(* IEC 61131-3 sources: STruCpp/tests/st-validation/oscat, 20 files *)

(* ---- oscat_bits.st ---- *)
FUNCTION BIT_TOGGLE_B : BYTE
VAR_INPUT
	IN : BYTE;
	POS : INT;
END_VAR
BIT_TOGGLE_B := SHL(BYTE#1, POS) XOR IN;
END_FUNCTION

FUNCTION BYTE_TO_GRAY : BYTE
VAR_INPUT
	IN : BYTE;
END_VAR
BYTE_TO_GRAY := IN XOR SHR(IN,1);
END_FUNCTION

FUNCTION GRAY_TO_BYTE : BYTE
VAR_INPUT
	IN : BYTE;
END_VAR
GRAY_TO_BYTE := SHR(IN,4) XOR IN;
GRAY_TO_BYTE := SHR(GRAY_TO_BYTE,2) XOR GRAY_TO_BYTE;
GRAY_TO_BYTE := SHR(GRAY_TO_BYTE,1) XOR GRAY_TO_BYTE;
END_FUNCTION

(* ---- oscat_convert.st ---- *)
(* OSCAT Conversion Functions — Unit conversions and range mapping *)

FUNCTION KMH_TO_MS : REAL
VAR_INPUT
	KMH : REAL;
END_VAR
KMH_TO_MS := KMH * 0.2777777777777;
END_FUNCTION

FUNCTION BFT_TO_MS : REAL
VAR_INPUT
	BFT : INT;
END_VAR
BFT_TO_MS := EXPT(BFT, 1.5) * 0.836;
END_FUNCTION

FUNCTION MS_TO_BFT : INT
VAR_INPUT
	MS : REAL;
END_VAR
MS_TO_BFT := REAL_TO_INT(EXPT(MS * 1.196172, 0.666667));
END_FUNCTION

FUNCTION BYTE_TO_RANGE : REAL
VAR_INPUT
	X : BYTE;
	LOW : REAL;
	HIGH : REAL;
END_VAR
BYTE_TO_RANGE := (HIGH - LOW) * X / 255.0 + LOW;
END_FUNCTION

FUNCTION RANGE_TO_BYTE : BYTE
VAR_INPUT
	X : REAL;
	LOW : REAL;
	HIGH : REAL;
END_VAR
RANGE_TO_BYTE := INT_TO_BYTE(TRUNC((LIMIT(LOW, X, HIGH) - LOW) * 255.0 / (HIGH - LOW)));
END_FUNCTION

(* ---- oscat_encoding.st ---- *)
(* OSCAT Encoding/Numeric Functions — BCD encoding and combinatorics *)

FUNCTION INT_TO_BCDC : BYTE
VAR_INPUT
	IN : INT;
END_VAR
INT_TO_BCDC := SHL(INT_TO_BYTE(IN / 10), 4) OR INT_TO_BYTE(IN MOD 10);
END_FUNCTION

FUNCTION BINOM : DINT
VAR_INPUT
	N : INT;
	K : INT;
END_VAR
VAR
	I : INT;
END_VAR
IF 2 * K > N THEN
	K := N - K;
END_IF;
IF K > N THEN
	RETURN;
ELSIF K = 0 OR K = N THEN
	BINOM := 1;
ELSIF K = 1 THEN
	BINOM := N;
ELSE
	BINOM := N;
	N := N + 1;
	FOR I := 2 TO K DO
		BINOM := BINOM * (N - I) / I;
	END_FOR;
END_IF;
END_FUNCTION

FUNCTION FIB : DINT
VAR_INPUT
	X : INT;
END_VAR
VAR
	T1 : DINT;
	T2 : DINT;
END_VAR
IF X < 0 OR X > 46 THEN
	FIB := -1;
ELSIF X < 2 THEN
	FIB := X;
	RETURN;
ELSE
	T2 := 1;
	WHILE X > 3 DO
		X := X - 2;
		T1 := T1 + T2;
		T2 := T1 + T2;
	END_WHILE;
	IF X > 2 THEN T1 := T1 + T2; END_IF;
	FIB := T1 + T2;
END_IF;
END_FUNCTION

(* ---- oscat_hyperbolic.st ---- *)
(* OSCAT Hyperbolic Math Functions — Pure math, no external dependencies *)

FUNCTION ACOSH : REAL
VAR_INPUT
	X : REAL;
END_VAR
ACOSH := LN(SQRT(X * X - 1.0) + X);
END_FUNCTION

FUNCTION ASINH : REAL
VAR_INPUT
	X : REAL;
END_VAR
ASINH := LN(SQRT(X * X + 1.0) + X);
END_FUNCTION

FUNCTION ATANH : REAL
VAR_INPUT
	X : REAL;
END_VAR
ATANH := LN((1.0 + X) / (1.0 - X)) * 0.5;
END_FUNCTION

FUNCTION ACOTH : REAL
VAR_INPUT
	X : REAL;
END_VAR
ACOTH := LN((X + 1.0) / (X - 1.0)) * 0.5;
END_FUNCTION

FUNCTION SIGN_R : BOOL
VAR_INPUT
	IN : REAL;
END_VAR
SIGN_R := IN < 0.0;
END_FUNCTION

(* ---- oscat_math.st ---- *)
FUNCTION MS_TO_KMH : REAL
VAR_INPUT
	ms : REAL;
END_VAR
MS_TO_KMH := ms * 3.6;
END_FUNCTION

FUNCTION NEGX : REAL
VAR_INPUT
	X : REAL;
END_VAR
NEGX := -X;
END_FUNCTION

FUNCTION HYPOT : REAL
VAR_INPUT
	X : REAL;
	Y : REAL;
END_VAR
HYPOT := SQRT(x*x + y*y);
END_FUNCTION

FUNCTION EXP10 : REAL
VAR_INPUT
	X : REAL;
END_VAR
EXP10 := EXP(X * 2.30258509299405);
END_FUNCTION

FUNCTION WINDOW : BOOL
VAR_INPUT
	low : REAL;
	in : REAL;
	high : REAL;
END_VAR
WINDOW := in < high AND in > low;
END_FUNCTION

FUNCTION WINDOW2 : BOOL
VAR_INPUT
	LOW : REAL;
	IN : REAL;
	HIGH : REAL;
END_VAR
WINDOW2 := IN >= LOW AND IN <= HIGH;
END_FUNCTION

FUNCTION SCALE : REAL
VAR_INPUT
	X : REAL;
	K : REAL;
	O : REAL;
	MX : REAL;
	MN : REAL;
END_VAR
SCALE := LIMIT(MN, X * K + O, MX);
END_FUNCTION

(* ---- oscat_string.st ---- *)
(* OSCAT String Functions — String manipulation using standard IEC string ops *)

FUNCTION TRIM : STRING(254)
VAR_INPUT
	STR : STRING(254);
END_VAR
VAR
	POS : INT;
END_VAR
TRIM := STR;
REPEAT
	POS := FIND(TRIM, ' ');
	IF POS > 0 THEN TRIM := REPLACE(TRIM, '', 1, POS); END_IF;
UNTIL POS = 0 END_REPEAT;
END_FUNCTION

FUNCTION TRIM1 : STRING(254)
VAR_INPUT
	STR : STRING(254);
END_VAR
VAR
	POS : INT;
END_VAR
TRIM1 := STR;
REPEAT
	POS := FIND(TRIM1, '  ');
	IF POS > 0 THEN TRIM1 := REPLACE(TRIM1, ' ', 2, POS); END_IF;
UNTIL POS = 0 END_REPEAT;
IF LEFT(TRIM1, 1) = ' ' THEN TRIM1 := DELETE(TRIM1, 1, 1); END_IF;
IF RIGHT(TRIM1, 1) = ' ' THEN TRIM1 := DELETE(TRIM1, 1, LEN(TRIM1)); END_IF;
END_FUNCTION

FUNCTION FINDB : INT
VAR_INPUT
	STR1 : STRING(254);
	STR2 : STRING(254);
END_VAR
VAR
	POS : INT;
	LENGTH : INT;
END_VAR
LENGTH := LEN(STR2);
FOR POS := LEN(STR1) - LENGTH + 1 TO 1 BY -1 DO
	IF MID(STR1, LENGTH, POS) = STR2 THEN
		FINDB := POS;
		RETURN;
	END_IF;
END_FOR;
FINDB := 0;
END_FUNCTION

FUNCTION REPLACE_CHARS : STRING(254)
VAR_INPUT
	STR : STRING(254);
	SRC : STRING(254);
	REP : STRING(254);
END_VAR
VAR
	A : INT;
	B : INT;
	C : STRING(1);
	STP : INT;
END_VAR
REPLACE_CHARS := STR;
A := LEN(SRC);
B := LEN(REP);
IF A < B THEN
	REP := LEFT(REP, A);
ELSIF B < A THEN
	SRC := LEFT(SRC, B);
END_IF;
STP := LEN(STR);
FOR A := 1 TO STP DO
	C := MID(REPLACE_CHARS, 1, A);
	B := FIND(SRC, C);
	IF B > 0 THEN
		REPLACE_CHARS := REPLACE(REPLACE_CHARS, MID(REP, 1, B), 1, A);
	END_IF;
END_FOR;
END_FUNCTION

(* ---- oscat_trig.st ---- *)
FUNCTION FLOOR2 : DINT
VAR_INPUT
	X : REAL;
END_VAR
FLOOR2 := REAL_TO_DINT(X);
IF DINT_TO_REAL(FLOOR2) > X THEN
	FLOOR2 := FLOOR2 - 1;
END_IF;
END_FUNCTION

FUNCTION MODR : REAL
VAR_INPUT
	IN : REAL;
	DIVI : REAL;
END_VAR
IF divi = 0.0 THEN
	MODR := 0.0;
ELSE
	MODR := in - DINT_TO_REAL(FLOOR2(in / divi)) * divi;
END_IF;
END_FUNCTION

FUNCTION DEG : REAL
VAR_INPUT
	rad : REAL;
END_VAR
DEG := MODR(57.29577951308232 * RAD, 360.0);
END_FUNCTION

(* ---- oscat_control.st ---- *)
(* OSCAT Control Function Blocks — Stateful control elements *)

FUNCTION_BLOCK TOGGLE
VAR_INPUT
	CLK : BOOL;
	RST : BOOL;
END_VAR
VAR_OUTPUT
	Q : BOOL;
END_VAR
VAR
	EDGE : BOOL;
END_VAR
IF RST THEN
	Q := FALSE;
ELSIF CLK AND NOT EDGE THEN
	Q := NOT Q;
END_IF;
EDGE := CLK;
END_FUNCTION_BLOCK

FUNCTION_BLOCK HYST_1
VAR_INPUT
	IN : REAL;
	HIGH : REAL;
	LOW : REAL;
END_VAR
VAR_OUTPUT
	Q : BOOL;
	WIN : BOOL;
END_VAR
IF IN < LOW THEN
	Q := FALSE;
	WIN := FALSE;
ELSIF IN > HIGH THEN
	Q := TRUE;
	WIN := FALSE;
ELSE
	WIN := TRUE;
END_IF;
END_FUNCTION_BLOCK

FUNCTION_BLOCK MANUAL_1
VAR_INPUT
	IN : BOOL;
	MAN : BOOL;
	M_I : BOOL;
	SET : BOOL;
	RST : BOOL;
END_VAR
VAR_OUTPUT
	Q : BOOL;
	STATUS : BYTE;
END_VAR
VAR
	S_EDGE : BOOL;
	R_EDGE : BOOL;
	MEDGE : BOOL;
END_VAR
IF NOT MAN THEN
	Q := IN;
	STATUS := 100;
	MEDGE := FALSE;
ELSIF NOT S_EDGE AND SET THEN
	Q := TRUE;
	MEDGE := TRUE;
	STATUS := 101;
ELSIF NOT R_EDGE AND RST THEN
	Q := FALSE;
	MEDGE := TRUE;
	STATUS := 102;
ELSIF NOT MEDGE THEN
	Q := M_I;
	STATUS := 103;
END_IF;
S_EDGE := SET;
R_EDGE := RST;
END_FUNCTION_BLOCK

(* ---- oscat_fb.st ---- *)
FUNCTION INC : INT
VAR_INPUT
	X : INT;
	D : INT;
	M : INT;
END_VAR
INC := (X + D + M + 1) MOD (M + 1);
END_FUNCTION

FUNCTION_BLOCK FF_DRE
VAR_INPUT
	SET : BOOL;
	D : BOOL;
	CLK : BOOL;
	RST : BOOL;
END_VAR
VAR_OUTPUT
	Q : BOOL;
END_VAR
VAR
	edge : BOOL;
END_VAR
IF rst OR set THEN
	Q := NOT rst;
ELSIF clk AND NOT edge THEN
	Q := D;
END_IF;
edge := CLK;
END_FUNCTION_BLOCK

FUNCTION_BLOCK COUNT_BR
VAR_INPUT
	SET : BOOL;
	IN : BYTE;
	UP : BOOL;
	DN : BOOL;
	STEP : BYTE := 1;
	MX : BYTE := 255;
	RST : BOOL;
END_VAR
VAR_OUTPUT
	CNT : BYTE;
END_VAR
VAR
	last_up: BOOL;
	last_dn: BOOL;
END_VAR
IF rst THEN
	cnt := 0;
ELSIF set THEN
	cnt := LIMIT(0,in,mx);
ELSIF up AND NOT last_up THEN
	cnt := INT_TO_BYTE(INC(cnt,step,mx));
ELSIF dn AND NOT last_dn THEN
	cnt := INT_TO_BYTE(inc(cnt,-step,mx));
END_IF;
last_up := up;
last_dn := dn;
END_FUNCTION_BLOCK

(* ---- oscat_logic.st ---- *)
(* OSCAT Logic Function Blocks — Flip-flops and sequential logic *)

FUNCTION_BLOCK FF_JKE
VAR_INPUT
	SET : BOOL;
	J : BOOL;
	CLK : BOOL;
	K : BOOL;
	RST : BOOL;
END_VAR
VAR_OUTPUT
	Q : BOOL;
END_VAR
VAR
	EDGE : BOOL;
END_VAR
IF RST OR SET THEN
	Q := NOT RST;
ELSIF CLK AND NOT EDGE THEN
	IF J XOR K THEN
		Q := J;
	ELSE
		Q := K XOR Q;
	END_IF;
END_IF;
EDGE := CLK;
END_FUNCTION_BLOCK

FUNCTION FLOOR2 : DINT
VAR_INPUT
	X : REAL;
END_VAR
FLOOR2 := REAL_TO_DINT(X);
IF DINT_TO_REAL(FLOOR2) > X THEN
	FLOOR2 := FLOOR2 - 1;
END_IF;
END_FUNCTION

FUNCTION MODR : REAL
VAR_INPUT
	IN : REAL;
	DIVI : REAL;
END_VAR
IF DIVI = 0.0 THEN
	MODR := 0.0;
ELSE
	MODR := IN - DINT_TO_REAL(FLOOR2(IN / DIVI)) * DIVI;
END_IF;
END_FUNCTION

(* ---- test_oscat_bits.st ---- *)
(* OSCAT Bit Manipulation Functions — End-to-End Tests *)

(* === BIT_TOGGLE_B: toggle a bit in a BYTE at a given position === *)

TEST 'BIT_TOGGLE_B: toggle bit 0 of 0 -> 1'
  VAR result : BYTE; END_VAR
  result := BIT_TOGGLE_B(IN := 0, POS := 0);
  ASSERT_EQ(result, 1);
END_TEST

TEST 'BIT_TOGGLE_B: toggle bit 0 of 1 -> 0'
  VAR result : BYTE; END_VAR
  result := BIT_TOGGLE_B(IN := 1, POS := 0);
  ASSERT_EQ(result, 0);
END_TEST

TEST 'BIT_TOGGLE_B: toggle bit 7 of 0 -> 128'
  VAR result : BYTE; END_VAR
  result := BIT_TOGGLE_B(IN := 0, POS := 7);
  ASSERT_EQ(result, 128);
END_TEST

TEST 'BIT_TOGGLE_B: toggle bit 3 of 255 -> 247'
  VAR result : BYTE; END_VAR
  result := BIT_TOGGLE_B(IN := 255, POS := 3);
  ASSERT_EQ(result, 247);
END_TEST

TEST 'BIT_TOGGLE_B: toggle bit 4 of 16#AA -> 16#BA'
  VAR result : BYTE; END_VAR
  result := BIT_TOGGLE_B(IN := 16#AA, POS := 4);
  (* 16#AA = 10101010, toggle bit 4 -> 10111010 = 16#BA = 186 *)
  ASSERT_EQ(result, 186);
END_TEST

(* === BYTE_TO_GRAY: binary to Gray code === *)

TEST 'BYTE_TO_GRAY: 0 -> 0'
  VAR result : BYTE; END_VAR
  result := BYTE_TO_GRAY(IN := 0);
  ASSERT_EQ(result, 0);
END_TEST

TEST 'BYTE_TO_GRAY: 1 -> 1'
  VAR result : BYTE; END_VAR
  result := BYTE_TO_GRAY(IN := 1);
  ASSERT_EQ(result, 1);
END_TEST

TEST 'BYTE_TO_GRAY: 2 -> 3'
  VAR result : BYTE; END_VAR
  result := BYTE_TO_GRAY(IN := 2);
  ASSERT_EQ(result, 3);
END_TEST

TEST 'BYTE_TO_GRAY: 3 -> 2'
  VAR result : BYTE; END_VAR
  result := BYTE_TO_GRAY(IN := 3);
  ASSERT_EQ(result, 2);
END_TEST

TEST 'BYTE_TO_GRAY: 4 -> 6'
  VAR result : BYTE; END_VAR
  result := BYTE_TO_GRAY(IN := 4);
  ASSERT_EQ(result, 6);
END_TEST

TEST 'BYTE_TO_GRAY: 255 -> 128'
  VAR result : BYTE; END_VAR
  result := BYTE_TO_GRAY(IN := 255);
  ASSERT_EQ(result, 128);
END_TEST

(* === GRAY_TO_BYTE: Gray code to binary === *)

TEST 'GRAY_TO_BYTE: 0 -> 0'
  VAR result : BYTE; END_VAR
  result := GRAY_TO_BYTE(IN := 0);
  ASSERT_EQ(result, 0);
END_TEST

TEST 'GRAY_TO_BYTE: 1 -> 1'
  VAR result : BYTE; END_VAR
  result := GRAY_TO_BYTE(IN := 1);
  ASSERT_EQ(result, 1);
END_TEST

TEST 'GRAY_TO_BYTE: 3 -> 2'
  VAR result : BYTE; END_VAR
  result := GRAY_TO_BYTE(IN := 3);
  ASSERT_EQ(result, 2);
END_TEST

TEST 'GRAY_TO_BYTE: 2 -> 3'
  VAR result : BYTE; END_VAR
  result := GRAY_TO_BYTE(IN := 2);
  ASSERT_EQ(result, 3);
END_TEST

TEST 'GRAY_TO_BYTE: 128 -> 255'
  VAR result : BYTE; END_VAR
  result := GRAY_TO_BYTE(IN := 128);
  ASSERT_EQ(result, 255);
END_TEST

(* === Round-trip: BYTE_TO_GRAY then GRAY_TO_BYTE === *)

TEST 'Round-trip: Gray(42) back to 42'
  VAR gray : BYTE; result : BYTE; END_VAR
  gray := BYTE_TO_GRAY(IN := 42);
  result := GRAY_TO_BYTE(IN := gray);
  ASSERT_EQ(result, 42);
END_TEST

TEST 'Round-trip: Gray(100) back to 100'
  VAR gray : BYTE; result : BYTE; END_VAR
  gray := BYTE_TO_GRAY(IN := 100);
  result := GRAY_TO_BYTE(IN := gray);
  ASSERT_EQ(result, 100);
END_TEST

TEST 'Round-trip: Gray(200) back to 200'
  VAR gray : BYTE; result : BYTE; END_VAR
  gray := BYTE_TO_GRAY(IN := 200);
  result := GRAY_TO_BYTE(IN := gray);
  ASSERT_EQ(result, 200);
END_TEST

(* ---- test_oscat_control.st ---- *)
(* OSCAT Control Function Blocks — End-to-End Tests *)

(* === TOGGLE: toggle output on rising clock edge === *)

TEST 'TOGGLE: initial Q is FALSE'
  VAR t : TOGGLE; END_VAR
  t(CLK := FALSE, RST := FALSE);
  ASSERT_FALSE(t.Q);
END_TEST

TEST 'TOGGLE: first rising edge toggles Q TRUE'
  VAR t : TOGGLE; END_VAR
  t(CLK := FALSE, RST := FALSE);
  t(CLK := TRUE, RST := FALSE);
  ASSERT_TRUE(t.Q);
END_TEST

TEST 'TOGGLE: second rising edge toggles Q FALSE'
  VAR t : TOGGLE; END_VAR
  t(CLK := FALSE, RST := FALSE);
  t(CLK := TRUE, RST := FALSE);
  ASSERT_TRUE(t.Q);
  t(CLK := FALSE, RST := FALSE);
  t(CLK := TRUE, RST := FALSE);
  ASSERT_FALSE(t.Q);
END_TEST

TEST 'TOGGLE: sustained CLK high does not toggle'
  VAR t : TOGGLE; END_VAR
  t(CLK := FALSE, RST := FALSE);
  t(CLK := TRUE, RST := FALSE);
  ASSERT_TRUE(t.Q);
  t(CLK := TRUE, RST := FALSE);
  ASSERT_TRUE(t.Q);
END_TEST

TEST 'TOGGLE: RST forces Q FALSE'
  VAR t : TOGGLE; END_VAR
  t(CLK := FALSE, RST := FALSE);
  t(CLK := TRUE, RST := FALSE);
  ASSERT_TRUE(t.Q);
  t(CLK := FALSE, RST := TRUE);
  ASSERT_FALSE(t.Q);
END_TEST

(* === HYST_1: simple hysteresis === *)

TEST 'HYST_1: below low -> Q FALSE'
  VAR h : HYST_1; END_VAR
  h(IN := 5.0, HIGH := 80.0, LOW := 20.0);
  ASSERT_FALSE(h.Q);
  ASSERT_FALSE(h.WIN);
END_TEST

TEST 'HYST_1: above high -> Q TRUE'
  VAR h : HYST_1; END_VAR
  h(IN := 90.0, HIGH := 80.0, LOW := 20.0);
  ASSERT_TRUE(h.Q);
  ASSERT_FALSE(h.WIN);
END_TEST

TEST 'HYST_1: in window -> WIN TRUE, Q unchanged'
  VAR h : HYST_1; END_VAR
  h(IN := 50.0, HIGH := 80.0, LOW := 20.0);
  ASSERT_TRUE(h.WIN);
END_TEST

TEST 'HYST_1: hysteresis holds Q through window'
  VAR h : HYST_1; END_VAR
  h(IN := 90.0, HIGH := 80.0, LOW := 20.0);
  ASSERT_TRUE(h.Q);
  h(IN := 50.0, HIGH := 80.0, LOW := 20.0);
  ASSERT_TRUE(h.Q);
  ASSERT_TRUE(h.WIN);
END_TEST

TEST 'HYST_1: crossing low clears Q'
  VAR h : HYST_1; END_VAR
  h(IN := 90.0, HIGH := 80.0, LOW := 20.0);
  ASSERT_TRUE(h.Q);
  h(IN := 10.0, HIGH := 80.0, LOW := 20.0);
  ASSERT_FALSE(h.Q);
END_TEST

(* === MANUAL_1: automatic/manual mode selector === *)

TEST 'MANUAL_1: auto mode passes IN to Q'
  VAR m : MANUAL_1; END_VAR
  m(IN := TRUE, MAN := FALSE, M_I := FALSE, SET := FALSE, RST := FALSE);
  ASSERT_TRUE(m.Q);
  ASSERT_EQ(m.STATUS, 100);
END_TEST

TEST 'MANUAL_1: auto mode with IN FALSE'
  VAR m : MANUAL_1; END_VAR
  m(IN := FALSE, MAN := FALSE, M_I := FALSE, SET := FALSE, RST := FALSE);
  ASSERT_FALSE(m.Q);
  ASSERT_EQ(m.STATUS, 100);
END_TEST

TEST 'MANUAL_1: manual SET forces Q TRUE'
  VAR m : MANUAL_1; END_VAR
  m(IN := FALSE, MAN := TRUE, M_I := FALSE, SET := FALSE, RST := FALSE);
  m(IN := FALSE, MAN := TRUE, M_I := FALSE, SET := TRUE, RST := FALSE);
  ASSERT_TRUE(m.Q);
  ASSERT_EQ(m.STATUS, 101);
END_TEST

TEST 'MANUAL_1: manual RST forces Q FALSE'
  VAR m : MANUAL_1; END_VAR
  m(IN := FALSE, MAN := TRUE, M_I := FALSE, SET := FALSE, RST := FALSE);
  m(IN := FALSE, MAN := TRUE, M_I := FALSE, SET := FALSE, RST := TRUE);
  ASSERT_FALSE(m.Q);
  ASSERT_EQ(m.STATUS, 102);
END_TEST

TEST 'MANUAL_1: manual M_I passthrough when no edges'
  VAR m : MANUAL_1; END_VAR
  m(IN := FALSE, MAN := TRUE, M_I := TRUE, SET := FALSE, RST := FALSE);
  ASSERT_TRUE(m.Q);
  ASSERT_EQ(m.STATUS, 103);
END_TEST

(* ---- test_oscat_convert.st ---- *)
(* OSCAT Conversion Functions — End-to-End Tests *)

(* === KMH_TO_MS: km/h to m/s === *)

TEST 'KMH_TO_MS: 3.6 km/h = 1 m/s'
  VAR result : REAL; END_VAR
  result := KMH_TO_MS(KMH := 3.6);
  ASSERT_NEAR(result, 1.0, 0.001);
END_TEST

TEST 'KMH_TO_MS: 100 km/h ~ 27.778 m/s'
  VAR result : REAL; END_VAR
  result := KMH_TO_MS(KMH := 100.0);
  ASSERT_NEAR(result, 27.778, 0.01);
END_TEST

TEST 'KMH_TO_MS: 0 km/h = 0 m/s'
  VAR result : REAL; END_VAR
  result := KMH_TO_MS(KMH := 0.0);
  ASSERT_NEAR(result, 0.0, 0.001);
END_TEST

(* === BFT_TO_MS: Beaufort to m/s === *)

TEST 'BFT_TO_MS: Beaufort 0 = 0 m/s'
  VAR result : REAL; END_VAR
  result := BFT_TO_MS(BFT := 0);
  ASSERT_NEAR(result, 0.0, 0.001);
END_TEST

TEST 'BFT_TO_MS: Beaufort 1 ~ 0.836 m/s'
  VAR result : REAL; END_VAR
  result := BFT_TO_MS(BFT := 1);
  ASSERT_NEAR(result, 0.836, 0.01);
END_TEST

TEST 'BFT_TO_MS: Beaufort 4 ~ 6.688 m/s'
  VAR result : REAL; END_VAR
  result := BFT_TO_MS(BFT := 4);
  ASSERT_NEAR(result, 6.688, 0.1);
END_TEST

(* === MS_TO_BFT: m/s to Beaufort === *)

TEST 'MS_TO_BFT: 0 m/s = Beaufort 0'
  VAR result : INT; END_VAR
  result := MS_TO_BFT(MS := 0.0);
  ASSERT_EQ(result, 0);
END_TEST

TEST 'MS_TO_BFT: 0.836 m/s ~ Beaufort 1'
  VAR result : INT; END_VAR
  result := MS_TO_BFT(MS := 0.836);
  ASSERT_EQ(result, 1);
END_TEST

(* === BYTE_TO_RANGE: byte to real range === *)

TEST 'BYTE_TO_RANGE: 0 maps to low'
  VAR result : REAL; END_VAR
  result := BYTE_TO_RANGE(X := 0, LOW := 0.0, HIGH := 100.0);
  ASSERT_NEAR(result, 0.0, 0.01);
END_TEST

TEST 'BYTE_TO_RANGE: 255 maps to high'
  VAR result : REAL; END_VAR
  result := BYTE_TO_RANGE(X := 255, LOW := 0.0, HIGH := 100.0);
  ASSERT_NEAR(result, 100.0, 0.01);
END_TEST

TEST 'BYTE_TO_RANGE: 127 maps to midpoint'
  VAR result : REAL; END_VAR
  result := BYTE_TO_RANGE(X := 127, LOW := 0.0, HIGH := 100.0);
  ASSERT_NEAR(result, 49.8, 0.2);
END_TEST

TEST 'BYTE_TO_RANGE: negative range'
  VAR result : REAL; END_VAR
  result := BYTE_TO_RANGE(X := 0, LOW := -10.0, HIGH := 10.0);
  ASSERT_NEAR(result, -10.0, 0.01);
END_TEST

(* === RANGE_TO_BYTE: real range to byte === *)

TEST 'RANGE_TO_BYTE: low maps to 0'
  VAR result : BYTE; END_VAR
  result := RANGE_TO_BYTE(X := 0.0, LOW := 0.0, HIGH := 100.0);
  ASSERT_EQ(result, 0);
END_TEST

TEST 'RANGE_TO_BYTE: high maps to 255'
  VAR result : BYTE; END_VAR
  result := RANGE_TO_BYTE(X := 100.0, LOW := 0.0, HIGH := 100.0);
  ASSERT_EQ(result, 255);
END_TEST

TEST 'RANGE_TO_BYTE: midpoint maps to ~127'
  VAR result : BYTE; END_VAR
  result := RANGE_TO_BYTE(X := 50.0, LOW := 0.0, HIGH := 100.0);
  ASSERT_EQ(result, 127);
END_TEST

TEST 'RANGE_TO_BYTE: clamps below to 0'
  VAR result : BYTE; END_VAR
  result := RANGE_TO_BYTE(X := -10.0, LOW := 0.0, HIGH := 100.0);
  ASSERT_EQ(result, 0);
END_TEST

TEST 'RANGE_TO_BYTE: clamps above to 255'
  VAR result : BYTE; END_VAR
  result := RANGE_TO_BYTE(X := 200.0, LOW := 0.0, HIGH := 100.0);
  ASSERT_EQ(result, 255);
END_TEST

(* ---- test_oscat_encoding.st ---- *)
(* OSCAT Encoding/Numeric Functions — End-to-End Tests *)

(* === INT_TO_BCDC: integer to BCD byte === *)

TEST 'INT_TO_BCDC: 0 -> 0x00'
  VAR result : BYTE; END_VAR
  result := INT_TO_BCDC(IN := 0);
  ASSERT_EQ(result, 0);
END_TEST

TEST 'INT_TO_BCDC: 9 -> 0x09'
  VAR result : BYTE; END_VAR
  result := INT_TO_BCDC(IN := 9);
  ASSERT_EQ(result, 9);
END_TEST

TEST 'INT_TO_BCDC: 10 -> 0x10'
  VAR result : BYTE; END_VAR
  result := INT_TO_BCDC(IN := 10);
  ASSERT_EQ(result, 16);
END_TEST

TEST 'INT_TO_BCDC: 42 -> 0x42'
  VAR result : BYTE; END_VAR
  result := INT_TO_BCDC(IN := 42);
  ASSERT_EQ(result, 66);
END_TEST

TEST 'INT_TO_BCDC: 99 -> 0x99'
  VAR result : BYTE; END_VAR
  result := INT_TO_BCDC(IN := 99);
  ASSERT_EQ(result, 153);
END_TEST

(* === BINOM: binomial coefficient C(n,k) === *)

TEST 'BINOM: C(0,0) = 1'
  VAR result : DINT; END_VAR
  result := BINOM(N := 0, K := 0);
  ASSERT_EQ(result, 1);
END_TEST

TEST 'BINOM: C(5,0) = 1'
  VAR result : DINT; END_VAR
  result := BINOM(N := 5, K := 0);
  ASSERT_EQ(result, 1);
END_TEST

TEST 'BINOM: C(5,1) = 5'
  VAR result : DINT; END_VAR
  result := BINOM(N := 5, K := 1);
  ASSERT_EQ(result, 5);
END_TEST

TEST 'BINOM: C(5,2) = 10'
  VAR result : DINT; END_VAR
  result := BINOM(N := 5, K := 2);
  ASSERT_EQ(result, 10);
END_TEST

TEST 'BINOM: C(10,3) = 120'
  VAR result : DINT; END_VAR
  result := BINOM(N := 10, K := 3);
  ASSERT_EQ(result, 120);
END_TEST

TEST 'BINOM: C(10,5) = 252'
  VAR result : DINT; END_VAR
  result := BINOM(N := 10, K := 5);
  ASSERT_EQ(result, 252);
END_TEST

TEST 'BINOM: C(20,10) = 184756'
  VAR result : DINT; END_VAR
  result := BINOM(N := 20, K := 10);
  ASSERT_EQ(result, 184756);
END_TEST

(* === FIB: Fibonacci number === *)

TEST 'FIB: fib(0) = 0'
  VAR result : DINT; END_VAR
  result := FIB(X := 0);
  ASSERT_EQ(result, 0);
END_TEST

TEST 'FIB: fib(1) = 1'
  VAR result : DINT; END_VAR
  result := FIB(X := 1);
  ASSERT_EQ(result, 1);
END_TEST

TEST 'FIB: fib(2) = 1'
  VAR result : DINT; END_VAR
  result := FIB(X := 2);
  ASSERT_EQ(result, 1);
END_TEST

TEST 'FIB: fib(5) = 5'
  VAR result : DINT; END_VAR
  result := FIB(X := 5);
  ASSERT_EQ(result, 5);
END_TEST

TEST 'FIB: fib(10) = 55'
  VAR result : DINT; END_VAR
  result := FIB(X := 10);
  ASSERT_EQ(result, 55);
END_TEST

TEST 'FIB: fib(20) = 6765'
  VAR result : DINT; END_VAR
  result := FIB(X := 20);
  ASSERT_EQ(result, 6765);
END_TEST

TEST 'FIB: negative input returns -1'
  VAR result : DINT; END_VAR
  result := FIB(X := -1);
  ASSERT_EQ(result, -1);
END_TEST

TEST 'FIB: overflow input returns -1'
  VAR result : DINT; END_VAR
  result := FIB(X := 47);
  ASSERT_EQ(result, -1);
END_TEST

(* ---- test_oscat_fb.st ---- *)
(* OSCAT Function Blocks — End-to-End Tests *)
(* Tests keyword identifiers (SET as VAR_INPUT) and FB state behavior *)

(* === FF_DRE: D-type flip-flop with rising edge clock === *)

TEST 'FF_DRE: initial state is FALSE'
  VAR ff : FF_DRE; END_VAR
  ff(SET := FALSE, D := FALSE, CLK := FALSE, RST := FALSE);
  ASSERT_FALSE(ff.Q);
END_TEST

TEST 'FF_DRE: SET forces Q TRUE'
  VAR ff : FF_DRE; END_VAR
  ff(SET := TRUE, D := FALSE, CLK := FALSE, RST := FALSE);
  ASSERT_TRUE(ff.Q);
END_TEST

TEST 'FF_DRE: RST forces Q FALSE'
  VAR ff : FF_DRE; END_VAR
  (* First set Q to TRUE *)
  ff(SET := TRUE, D := FALSE, CLK := FALSE, RST := FALSE);
  ASSERT_TRUE(ff.Q);
  (* Then reset *)
  ff(SET := FALSE, D := FALSE, CLK := FALSE, RST := TRUE);
  ASSERT_FALSE(ff.Q);
END_TEST

TEST 'FF_DRE: RST overrides SET'
  VAR ff : FF_DRE; END_VAR
  ff(SET := TRUE, D := TRUE, CLK := FALSE, RST := TRUE);
  ASSERT_FALSE(ff.Q);
END_TEST

TEST 'FF_DRE: rising CLK edge captures D=TRUE'
  VAR ff : FF_DRE; END_VAR
  (* CLK low first to establish edge *)
  ff(SET := FALSE, D := TRUE, CLK := FALSE, RST := FALSE);
  ASSERT_FALSE(ff.Q);
  (* Rising edge with D=TRUE *)
  ff(SET := FALSE, D := TRUE, CLK := TRUE, RST := FALSE);
  ASSERT_TRUE(ff.Q);
END_TEST

TEST 'FF_DRE: rising CLK edge captures D=FALSE'
  VAR ff : FF_DRE; END_VAR
  (* First set Q high *)
  ff(SET := TRUE, D := FALSE, CLK := FALSE, RST := FALSE);
  ASSERT_TRUE(ff.Q);
  (* CLK low to prepare edge *)
  ff(SET := FALSE, D := FALSE, CLK := FALSE, RST := FALSE);
  (* Rising edge with D=FALSE *)
  ff(SET := FALSE, D := FALSE, CLK := TRUE, RST := FALSE);
  ASSERT_FALSE(ff.Q);
END_TEST

TEST 'FF_DRE: no change on sustained CLK high'
  VAR ff : FF_DRE; END_VAR
  (* Rising edge captures D=TRUE *)
  ff(SET := FALSE, D := TRUE, CLK := FALSE, RST := FALSE);
  ff(SET := FALSE, D := TRUE, CLK := TRUE, RST := FALSE);
  ASSERT_TRUE(ff.Q);
  (* Now D changes but CLK stays high — no edge, no capture *)
  ff(SET := FALSE, D := FALSE, CLK := TRUE, RST := FALSE);
  ASSERT_TRUE(ff.Q);
END_TEST

(* === COUNT_BR: byte counter with SET keyword input === *)

TEST 'COUNT_BR: initial count is 0'
  VAR ctr : COUNT_BR; END_VAR
  ctr(SET := FALSE, IN := 0, UP := FALSE, DN := FALSE, RST := FALSE);
  ASSERT_EQ(ctr.CNT, 0);
END_TEST

TEST 'COUNT_BR: RST resets count to 0'
  VAR ctr : COUNT_BR; END_VAR
  (* Count up once *)
  ctr(SET := FALSE, IN := 0, UP := FALSE, DN := FALSE, RST := FALSE);
  ctr(SET := FALSE, IN := 0, UP := TRUE, DN := FALSE, RST := FALSE);
  (* Now reset *)
  ctr(SET := FALSE, IN := 0, UP := FALSE, DN := FALSE, RST := TRUE);
  ASSERT_EQ(ctr.CNT, 0);
END_TEST

TEST 'COUNT_BR: SET loads IN value'
  VAR ctr : COUNT_BR; END_VAR
  ctr(SET := TRUE, IN := 42, UP := FALSE, DN := FALSE, MX := 255, RST := FALSE);
  ASSERT_EQ(ctr.CNT, 42);
END_TEST

TEST 'COUNT_BR: SET clamps IN to MX'
  VAR ctr : COUNT_BR; END_VAR
  ctr(SET := TRUE, IN := 200, UP := FALSE, DN := FALSE, MX := 100, RST := FALSE);
  ASSERT_EQ(ctr.CNT, 100);
END_TEST

TEST 'COUNT_BR: count up on rising edge'
  VAR ctr : COUNT_BR; END_VAR
  (* UP low *)
  ctr(SET := FALSE, IN := 0, UP := FALSE, DN := FALSE, STEP := 1, MX := 255, RST := FALSE);
  ASSERT_EQ(ctr.CNT, 0);
  (* UP rising edge *)
  ctr(SET := FALSE, IN := 0, UP := TRUE, DN := FALSE, STEP := 1, MX := 255, RST := FALSE);
  ASSERT_EQ(ctr.CNT, 1);
END_TEST

TEST 'COUNT_BR: count up multiple steps'
  VAR ctr : COUNT_BR; END_VAR
  ctr(SET := FALSE, IN := 0, UP := FALSE, DN := FALSE, STEP := 5, MX := 255, RST := FALSE);
  (* First rising edge: 0 + 5 = 5 *)
  ctr(SET := FALSE, IN := 0, UP := TRUE, DN := FALSE, STEP := 5, MX := 255, RST := FALSE);
  ASSERT_EQ(ctr.CNT, 5);
  (* Need falling edge before next count *)
  ctr(SET := FALSE, IN := 0, UP := FALSE, DN := FALSE, STEP := 5, MX := 255, RST := FALSE);
  (* Second rising edge: 5 + 5 = 10 *)
  ctr(SET := FALSE, IN := 0, UP := TRUE, DN := FALSE, STEP := 5, MX := 255, RST := FALSE);
  ASSERT_EQ(ctr.CNT, 10);
END_TEST

(* ---- test_oscat_hyperbolic.st ---- *)
(* OSCAT Hyperbolic Functions — End-to-End Tests *)

(* === ACOSH: inverse hyperbolic cosine === *)

TEST 'ACOSH: acosh(1) = 0'
  VAR result : REAL; END_VAR
  result := ACOSH(X := 1.0);
  ASSERT_NEAR(result, 0.0, 0.001);
END_TEST

TEST 'ACOSH: acosh(2) ~ 1.3169'
  VAR result : REAL; END_VAR
  result := ACOSH(X := 2.0);
  ASSERT_NEAR(result, 1.3169, 0.001);
END_TEST

TEST 'ACOSH: acosh(10) ~ 2.9932'
  VAR result : REAL; END_VAR
  result := ACOSH(X := 10.0);
  ASSERT_NEAR(result, 2.9932, 0.001);
END_TEST

(* === ASINH: inverse hyperbolic sine === *)

TEST 'ASINH: asinh(0) = 0'
  VAR result : REAL; END_VAR
  result := ASINH(X := 0.0);
  ASSERT_NEAR(result, 0.0, 0.001);
END_TEST

TEST 'ASINH: asinh(1) ~ 0.8814'
  VAR result : REAL; END_VAR
  result := ASINH(X := 1.0);
  ASSERT_NEAR(result, 0.8814, 0.001);
END_TEST

TEST 'ASINH: asinh(-1) ~ -0.8814'
  VAR result : REAL; END_VAR
  result := ASINH(X := -1.0);
  ASSERT_NEAR(result, -0.8814, 0.001);
END_TEST

TEST 'ASINH: asinh(5) ~ 2.3124'
  VAR result : REAL; END_VAR
  result := ASINH(X := 5.0);
  ASSERT_NEAR(result, 2.3124, 0.001);
END_TEST

(* === ATANH: inverse hyperbolic tangent === *)

TEST 'ATANH: atanh(0) = 0'
  VAR result : REAL; END_VAR
  result := ATANH(X := 0.0);
  ASSERT_NEAR(result, 0.0, 0.001);
END_TEST

TEST 'ATANH: atanh(0.5) ~ 0.5493'
  VAR result : REAL; END_VAR
  result := ATANH(X := 0.5);
  ASSERT_NEAR(result, 0.5493, 0.001);
END_TEST

TEST 'ATANH: atanh(-0.5) ~ -0.5493'
  VAR result : REAL; END_VAR
  result := ATANH(X := -0.5);
  ASSERT_NEAR(result, -0.5493, 0.001);
END_TEST

(* === ACOTH: inverse hyperbolic cotangent === *)

TEST 'ACOTH: acoth(2) ~ 0.5493'
  VAR result : REAL; END_VAR
  result := ACOTH(X := 2.0);
  ASSERT_NEAR(result, 0.5493, 0.001);
END_TEST

TEST 'ACOTH: acoth(5) ~ 0.2027'
  VAR result : REAL; END_VAR
  result := ACOTH(X := 5.0);
  ASSERT_NEAR(result, 0.2027, 0.001);
END_TEST

TEST 'ACOTH: acoth(-2) ~ -0.5493'
  VAR result : REAL; END_VAR
  result := ACOTH(X := -2.0);
  ASSERT_NEAR(result, -0.5493, 0.001);
END_TEST

(* === SIGN_R: returns TRUE if input is negative === *)

TEST 'SIGN_R: positive is FALSE'
  VAR result : BOOL; END_VAR
  result := SIGN_R(IN := 5.0);
  ASSERT_FALSE(result);
END_TEST

TEST 'SIGN_R: negative is TRUE'
  VAR result : BOOL; END_VAR
  result := SIGN_R(IN := -3.14);
  ASSERT_TRUE(result);
END_TEST

TEST 'SIGN_R: zero is FALSE'
  VAR result : BOOL; END_VAR
  result := SIGN_R(IN := 0.0);
  ASSERT_FALSE(result);
END_TEST

(* ---- test_oscat_logic.st ---- *)
(* OSCAT Logic Functions — End-to-End Tests *)

(* === FF_JKE: JK flip-flop with edge detection === *)

TEST 'FF_JKE: initial state is FALSE'
  VAR ff : FF_JKE; END_VAR
  ff(SET := FALSE, J := FALSE, CLK := FALSE, K := FALSE, RST := FALSE);
  ASSERT_FALSE(ff.Q);
END_TEST

TEST 'FF_JKE: SET forces Q TRUE'
  VAR ff : FF_JKE; END_VAR
  ff(SET := TRUE, J := FALSE, CLK := FALSE, K := FALSE, RST := FALSE);
  ASSERT_TRUE(ff.Q);
END_TEST

TEST 'FF_JKE: RST forces Q FALSE'
  VAR ff : FF_JKE; END_VAR
  ff(SET := TRUE, J := FALSE, CLK := FALSE, K := FALSE, RST := FALSE);
  ASSERT_TRUE(ff.Q);
  ff(SET := FALSE, J := FALSE, CLK := FALSE, K := FALSE, RST := TRUE);
  ASSERT_FALSE(ff.Q);
END_TEST

TEST 'FF_JKE: RST overrides SET'
  VAR ff : FF_JKE; END_VAR
  ff(SET := TRUE, J := FALSE, CLK := FALSE, K := FALSE, RST := TRUE);
  ASSERT_FALSE(ff.Q);
END_TEST

TEST 'FF_JKE: J=1 K=0 sets Q on rising edge'
  VAR ff : FF_JKE; END_VAR
  ff(SET := FALSE, J := TRUE, CLK := FALSE, K := FALSE, RST := FALSE);
  ff(SET := FALSE, J := TRUE, CLK := TRUE, K := FALSE, RST := FALSE);
  ASSERT_TRUE(ff.Q);
END_TEST

TEST 'FF_JKE: J=0 K=1 clears Q on rising edge'
  VAR ff : FF_JKE; END_VAR
  ff(SET := TRUE, J := FALSE, CLK := FALSE, K := FALSE, RST := FALSE);
  ASSERT_TRUE(ff.Q);
  ff(SET := FALSE, J := FALSE, CLK := FALSE, K := TRUE, RST := FALSE);
  ff(SET := FALSE, J := FALSE, CLK := TRUE, K := TRUE, RST := FALSE);
  ASSERT_FALSE(ff.Q);
END_TEST

TEST 'FF_JKE: J=1 K=1 toggles Q on rising edge'
  VAR ff : FF_JKE; END_VAR
  ff(SET := FALSE, J := TRUE, CLK := FALSE, K := TRUE, RST := FALSE);
  ASSERT_FALSE(ff.Q);
  ff(SET := FALSE, J := TRUE, CLK := TRUE, K := TRUE, RST := FALSE);
  ASSERT_TRUE(ff.Q);
  ff(SET := FALSE, J := TRUE, CLK := FALSE, K := TRUE, RST := FALSE);
  ff(SET := FALSE, J := TRUE, CLK := TRUE, K := TRUE, RST := FALSE);
  ASSERT_FALSE(ff.Q);
END_TEST

TEST 'FF_JKE: J=0 K=0 holds Q on rising edge'
  VAR ff : FF_JKE; END_VAR
  ff(SET := TRUE, J := FALSE, CLK := FALSE, K := FALSE, RST := FALSE);
  ASSERT_TRUE(ff.Q);
  ff(SET := FALSE, J := FALSE, CLK := FALSE, K := FALSE, RST := FALSE);
  ff(SET := FALSE, J := FALSE, CLK := TRUE, K := FALSE, RST := FALSE);
  ASSERT_TRUE(ff.Q);
END_TEST

(* === FLOOR2: floor function for REAL === *)

TEST 'FLOOR2: positive exact'
  VAR result : DINT; END_VAR
  result := FLOOR2(X := 3.0);
  ASSERT_EQ(result, 3);
END_TEST

TEST 'FLOOR2: positive fractional'
  VAR result : DINT; END_VAR
  result := FLOOR2(X := 3.99);
  ASSERT_EQ(result, 3);
END_TEST

TEST 'FLOOR2: negative fractional rounds down'
  VAR result : DINT; END_VAR
  result := FLOOR2(X := -3.14);
  ASSERT_EQ(result, -4);
END_TEST

(* === MODR: real modulo via FLOOR2 === *)

TEST 'MODR: 5.5 mod 2.5 = 0.5'
  VAR result : REAL; END_VAR
  result := MODR(IN := 5.5, DIVI := 2.5);
  ASSERT_NEAR(result, 0.5, 0.001);
END_TEST

TEST 'MODR: 10.0 mod 3.0 = 1.0'
  VAR result : REAL; END_VAR
  result := MODR(IN := 10.0, DIVI := 3.0);
  ASSERT_NEAR(result, 1.0, 0.001);
END_TEST

TEST 'MODR: division by 0 returns 0'
  VAR result : REAL; END_VAR
  result := MODR(IN := 5.0, DIVI := 0.0);
  ASSERT_NEAR(result, 0.0, 0.001);
END_TEST

(* ---- test_oscat_math.st ---- *)
(* OSCAT Math Functions — End-to-End Tests *)

(* === MS_TO_KMH: meters/second to km/h === *)

TEST 'MS_TO_KMH: 1 m/s = 3.6 km/h'
  VAR result : REAL; END_VAR
  result := MS_TO_KMH(ms := 1.0);
  ASSERT_NEAR(result, 3.6, 0.001);
END_TEST

TEST 'MS_TO_KMH: 0 m/s = 0 km/h'
  VAR result : REAL; END_VAR
  result := MS_TO_KMH(ms := 0.0);
  ASSERT_NEAR(result, 0.0, 0.001);
END_TEST

TEST 'MS_TO_KMH: 27.778 m/s ~ 100 km/h'
  VAR result : REAL; END_VAR
  result := MS_TO_KMH(ms := 27.778);
  ASSERT_NEAR(result, 100.0, 0.1);
END_TEST

(* === NEGX: negate real === *)

TEST 'NEGX: positive becomes negative'
  VAR result : REAL; END_VAR
  result := NEGX(X := 5.0);
  ASSERT_NEAR(result, -5.0, 0.001);
END_TEST

TEST 'NEGX: negative becomes positive'
  VAR result : REAL; END_VAR
  result := NEGX(X := -3.14);
  ASSERT_NEAR(result, 3.14, 0.001);
END_TEST

TEST 'NEGX: zero stays zero'
  VAR result : REAL; END_VAR
  result := NEGX(X := 0.0);
  ASSERT_NEAR(result, 0.0, 0.001);
END_TEST

(* === HYPOT: Pythagorean theorem === *)

TEST 'HYPOT: 3-4-5 triangle'
  VAR result : REAL; END_VAR
  result := HYPOT(X := 3.0, Y := 4.0);
  ASSERT_NEAR(result, 5.0, 0.001);
END_TEST

TEST 'HYPOT: unit vector'
  VAR result : REAL; END_VAR
  result := HYPOT(X := 1.0, Y := 0.0);
  ASSERT_NEAR(result, 1.0, 0.001);
END_TEST

TEST 'HYPOT: zero inputs'
  VAR result : REAL; END_VAR
  result := HYPOT(X := 0.0, Y := 0.0);
  ASSERT_NEAR(result, 0.0, 0.001);
END_TEST

TEST 'HYPOT: negative inputs'
  VAR result : REAL; END_VAR
  result := HYPOT(X := -3.0, Y := -4.0);
  ASSERT_NEAR(result, 5.0, 0.001);
END_TEST

(* === EXP10: 10^x === *)

TEST 'EXP10: 10^0 = 1'
  VAR result : REAL; END_VAR
  result := EXP10(X := 0.0);
  ASSERT_NEAR(result, 1.0, 0.001);
END_TEST

TEST 'EXP10: 10^1 = 10'
  VAR result : REAL; END_VAR
  result := EXP10(X := 1.0);
  ASSERT_NEAR(result, 10.0, 0.01);
END_TEST

TEST 'EXP10: 10^3 = 1000'
  VAR result : REAL; END_VAR
  result := EXP10(X := 3.0);
  ASSERT_NEAR(result, 1000.0, 1.0);
END_TEST

TEST 'EXP10: 10^-1 = 0.1'
  VAR result : REAL; END_VAR
  result := EXP10(X := -1.0);
  ASSERT_NEAR(result, 0.1, 0.001);
END_TEST

(* === WINDOW: open interval check === *)

TEST 'WINDOW: value inside range'
  VAR result : BOOL; END_VAR
  result := WINDOW(low := 0.0, in := 5.0, high := 10.0);
  ASSERT_TRUE(result);
END_TEST

TEST 'WINDOW: value below range'
  VAR result : BOOL; END_VAR
  result := WINDOW(low := 0.0, in := -1.0, high := 10.0);
  ASSERT_FALSE(result);
END_TEST

TEST 'WINDOW: value above range'
  VAR result : BOOL; END_VAR
  result := WINDOW(low := 0.0, in := 11.0, high := 10.0);
  ASSERT_FALSE(result);
END_TEST

TEST 'WINDOW: value at lower boundary is excluded'
  VAR result : BOOL; END_VAR
  result := WINDOW(low := 0.0, in := 0.0, high := 10.0);
  ASSERT_FALSE(result);
END_TEST

TEST 'WINDOW: value at upper boundary is excluded'
  VAR result : BOOL; END_VAR
  result := WINDOW(low := 0.0, in := 10.0, high := 10.0);
  ASSERT_FALSE(result);
END_TEST

(* === WINDOW2: closed interval check === *)

TEST 'WINDOW2: value inside range'
  VAR result : BOOL; END_VAR
  result := WINDOW2(LOW := 0.0, IN := 5.0, HIGH := 10.0);
  ASSERT_TRUE(result);
END_TEST

TEST 'WINDOW2: value at lower boundary is included'
  VAR result : BOOL; END_VAR
  result := WINDOW2(LOW := 0.0, IN := 0.0, HIGH := 10.0);
  ASSERT_TRUE(result);
END_TEST

TEST 'WINDOW2: value at upper boundary is included'
  VAR result : BOOL; END_VAR
  result := WINDOW2(LOW := 0.0, IN := 10.0, HIGH := 10.0);
  ASSERT_TRUE(result);
END_TEST

TEST 'WINDOW2: value below range'
  VAR result : BOOL; END_VAR
  result := WINDOW2(LOW := 0.0, IN := -0.001, HIGH := 10.0);
  ASSERT_FALSE(result);
END_TEST

(* === SCALE: linear scaling with limits === *)

TEST 'SCALE: identity with no offset'
  VAR result : REAL; END_VAR
  result := SCALE(X := 5.0, K := 1.0, O := 0.0, MX := 100.0, MN := 0.0);
  ASSERT_NEAR(result, 5.0, 0.001);
END_TEST

TEST 'SCALE: double with offset'
  VAR result : REAL; END_VAR
  result := SCALE(X := 3.0, K := 2.0, O := 10.0, MX := 100.0, MN := 0.0);
  ASSERT_NEAR(result, 16.0, 0.001);
END_TEST

TEST 'SCALE: clamp to max'
  VAR result : REAL; END_VAR
  result := SCALE(X := 100.0, K := 2.0, O := 0.0, MX := 50.0, MN := 0.0);
  ASSERT_NEAR(result, 50.0, 0.001);
END_TEST

TEST 'SCALE: clamp to min'
  VAR result : REAL; END_VAR
  result := SCALE(X := -100.0, K := 1.0, O := 0.0, MX := 50.0, MN := -10.0);
  ASSERT_NEAR(result, -10.0, 0.001);
END_TEST

(* ---- test_oscat_string.st ---- *)
(* OSCAT String Functions — End-to-End Tests *)

(* === TRIM: remove all spaces === *)

TEST 'TRIM: removes all spaces'
  VAR result : STRING(254); END_VAR
  result := TRIM(STR := 'hello world');
  ASSERT_EQ(result, 'helloworld');
END_TEST

TEST 'TRIM: no spaces unchanged'
  VAR result : STRING(254); END_VAR
  result := TRIM(STR := 'hello');
  ASSERT_EQ(result, 'hello');
END_TEST

TEST 'TRIM: leading and trailing spaces'
  VAR result : STRING(254); END_VAR
  result := TRIM(STR := ' hello ');
  ASSERT_EQ(result, 'hello');
END_TEST

TEST 'TRIM: all spaces becomes empty'
  VAR result : STRING(254); END_VAR
  result := TRIM(STR := '   ');
  ASSERT_EQ(result, '');
END_TEST

(* === TRIM1: collapse multiple spaces to single, strip leading/trailing === *)

TEST 'TRIM1: collapses double spaces'
  VAR result : STRING(254); END_VAR
  result := TRIM1(STR := 'hello  world');
  ASSERT_EQ(result, 'hello world');
END_TEST

TEST 'TRIM1: strips leading space'
  VAR result : STRING(254); END_VAR
  result := TRIM1(STR := ' hello');
  ASSERT_EQ(result, 'hello');
END_TEST

TEST 'TRIM1: strips trailing space'
  VAR result : STRING(254); END_VAR
  result := TRIM1(STR := 'hello ');
  ASSERT_EQ(result, 'hello');
END_TEST

TEST 'TRIM1: normalizes multiple spaces'
  VAR result : STRING(254); END_VAR
  result := TRIM1(STR := '  a   b  c  ');
  ASSERT_EQ(result, 'a b c');
END_TEST

(* === FINDB: find substring from end === *)

TEST 'FINDB: finds last occurrence'
  VAR result : INT; END_VAR
  result := FINDB(STR1 := 'abcabc', STR2 := 'abc');
  ASSERT_EQ(result, 4);
END_TEST

TEST 'FINDB: finds only occurrence'
  VAR result : INT; END_VAR
  result := FINDB(STR1 := 'hello', STR2 := 'ell');
  ASSERT_EQ(result, 2);
END_TEST

TEST 'FINDB: not found returns 0'
  VAR result : INT; END_VAR
  result := FINDB(STR1 := 'hello', STR2 := 'xyz');
  ASSERT_EQ(result, 0);
END_TEST

TEST 'FINDB: empty search string'
  VAR result : INT; END_VAR
  result := FINDB(STR1 := 'hello', STR2 := '');
  (* Empty substring: loop runs from LEN+1 down to 1, MID of length 0 = '' = str2 at pos LEN+1 *)
  ASSERT_EQ(result, 6);
END_TEST

(* === REPLACE_CHARS: character-by-character replacement === *)

TEST 'REPLACE_CHARS: single char replacement'
  VAR result : STRING(254); END_VAR
  result := REPLACE_CHARS(STR := 'hello', SRC := 'l', REP := 'r');
  ASSERT_EQ(result, 'herro');
END_TEST

TEST 'REPLACE_CHARS: multi char mapping'
  VAR result : STRING(254); END_VAR
  result := REPLACE_CHARS(STR := 'abc', SRC := 'abc', REP := 'xyz');
  ASSERT_EQ(result, 'xyz');
END_TEST

TEST 'REPLACE_CHARS: no matches unchanged'
  VAR result : STRING(254); END_VAR
  result := REPLACE_CHARS(STR := 'hello', SRC := 'xyz', REP := 'abc');
  ASSERT_EQ(result, 'hello');
END_TEST

(* ---- test_oscat_trig.st ---- *)
(* OSCAT Trigonometric/Math Functions with Dependencies *)
(* Tests multi-function call chains: DEG -> MODR -> FLOOR2 *)

(* === FLOOR2: floor function for REAL === *)

TEST 'FLOOR2: positive exact'
  VAR result : DINT; END_VAR
  result := FLOOR2(X := 3.0);
  ASSERT_EQ(result, 3);
END_TEST

TEST 'FLOOR2: positive fractional'
  VAR result : DINT; END_VAR
  result := FLOOR2(X := 3.14);
  ASSERT_EQ(result, 3);
END_TEST

TEST 'FLOOR2: negative fractional rounds down'
  VAR result : DINT; END_VAR
  result := FLOOR2(X := -3.14);
  ASSERT_EQ(result, -4);
END_TEST

TEST 'FLOOR2: zero'
  VAR result : DINT; END_VAR
  result := FLOOR2(X := 0.0);
  ASSERT_EQ(result, 0);
END_TEST

(* === MODR: real modulo === *)

TEST 'MODR: 5.5 mod 2.5 = 0.5'
  VAR result : REAL; END_VAR
  result := MODR(IN := 5.5, DIVI := 2.5);
  ASSERT_NEAR(result, 0.5, 0.001);
END_TEST

TEST 'MODR: 10.0 mod 3.0 = 1.0'
  VAR result : REAL; END_VAR
  result := MODR(IN := 10.0, DIVI := 3.0);
  ASSERT_NEAR(result, 1.0, 0.001);
END_TEST

TEST 'MODR: division by 0 returns 0'
  VAR result : REAL; END_VAR
  result := MODR(IN := 5.0, DIVI := 0.0);
  ASSERT_NEAR(result, 0.0, 0.001);
END_TEST

TEST 'MODR: exact multiple returns 0'
  VAR result : REAL; END_VAR
  result := MODR(IN := 6.0, DIVI := 3.0);
  ASSERT_NEAR(result, 0.0, 0.001);
END_TEST

(* === DEG: radians to degrees === *)

TEST 'DEG: 0 radians = 0 degrees'
  VAR result : REAL; END_VAR
  result := DEG(rad := 0.0);
  ASSERT_NEAR(result, 0.0, 0.01);
END_TEST

TEST 'DEG: PI radians ~ 180 degrees'
  VAR result : REAL; END_VAR
  result := DEG(rad := 3.14159265358979);
  ASSERT_NEAR(result, 180.0, 0.01);
END_TEST

TEST 'DEG: PI/2 radians ~ 90 degrees'
  VAR result : REAL; END_VAR
  result := DEG(rad := 1.5707963267949);
  ASSERT_NEAR(result, 90.0, 0.01);
END_TEST

TEST 'DEG: 2*PI radians wraps to 0 degrees'
  VAR result : REAL; END_VAR
  result := DEG(rad := 6.28318530717959);
  ASSERT_NEAR(result, 0.0, 0.1);
END_TEST

TEST 'DEG: negative radians wrap correctly'
  VAR result : REAL; END_VAR
  result := DEG(rad := -1.5707963267949);
  (* -90 degrees, modulo 360 should wrap *)
  ASSERT_NEAR(result, 270.0, 0.1);
END_TEST
